// TIA Portal V20 export
DATA_BLOCK "iDB_CamManual"   // DB9
// stored: InstanceOfName FB_CamManual, InstanceOfType FB
"FB_CamManual"
   // VAR_INPUT
   //    xManEtiketa : Bool;
   //    xManFolie : Bool;
   //    tLightDelay : Time;
   //    tTrigPulse : Time;
   // END_VAR
   // VAR
   //    tonEt : TON_TIME;
   //    tpEt { S7_SetPoint := 'True'} : TP_TIME;
   //    tonFo { S7_SetPoint := 'True'} : TON_TIME;
   //    tpFo { S7_SetPoint := 'True'} : TP_TIME;
   // END_VAR
BEGIN
END_DATA_BLOCK
